// SIMATIC S7-200 project (STEP 7-Micro/WIN), CPU 224XP CN REL 02.01

SYMBOL_TABLE USUARIO1
C_1              VD100
C_0              VD110
y_k              VD180
r_k              VD190
u_k              VD120
xh1_k_1          VD130
xh1_k            VD140
xh2_k_1          VD300
xh2_k            VD160
xh3_k_1          VD170
xh3_k            VD200
xp1_k            VD210    // X1_v
xp2_k            VD220    // X2_v
xp3_k            VD230    // X3_v
Ao               VD310
Bo               VD320
Co               VD330
Do               VD340
Eo               VD350
Fo               VD360
Go               VD370
Ho               VD380
Io               VD390
Jo               VD400
L1o              VD410
L2o              VD420
L3o              VD430
e_k              VD270
Ee               VD240
r_k_1            VD250
u_k_1            VD150
k1o              VD440
k2o              VD450
k3o              VD460
END_SYMBOL_TABLE

ORGANIZATION_BLOCK PRINCIPAL:OB1
TITLE=COMENTARIOS DEL PROGRAMA
BEGIN
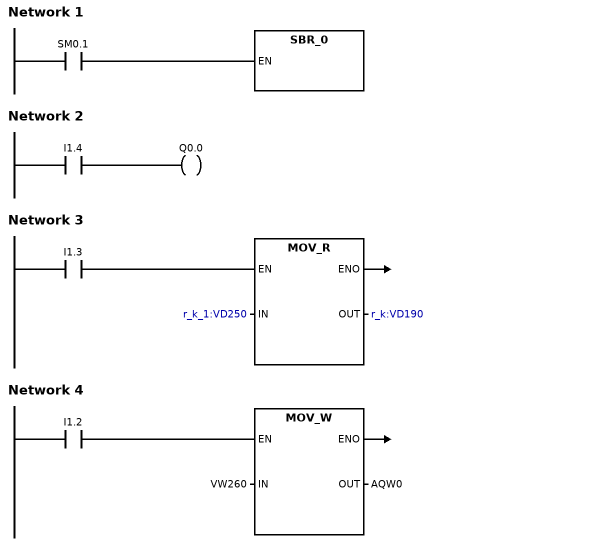
Network 1
LD     SM0.1
CALL   SBR_0:SBR0
Network 2
LD     I1.4
=      Q0.0
Network 3
LD     I1.3
MOVR   r_k_1:VD250, r_k:VD190
Network 4
LD     I1.2
MOVW   VW260, AQW0
END_ORGANIZATION_BLOCK

SUBROUTINE_BLOCK SBR_0:SBR0
TITLE=COMENTARIOS DE LA SUBRUTINA
BEGIN
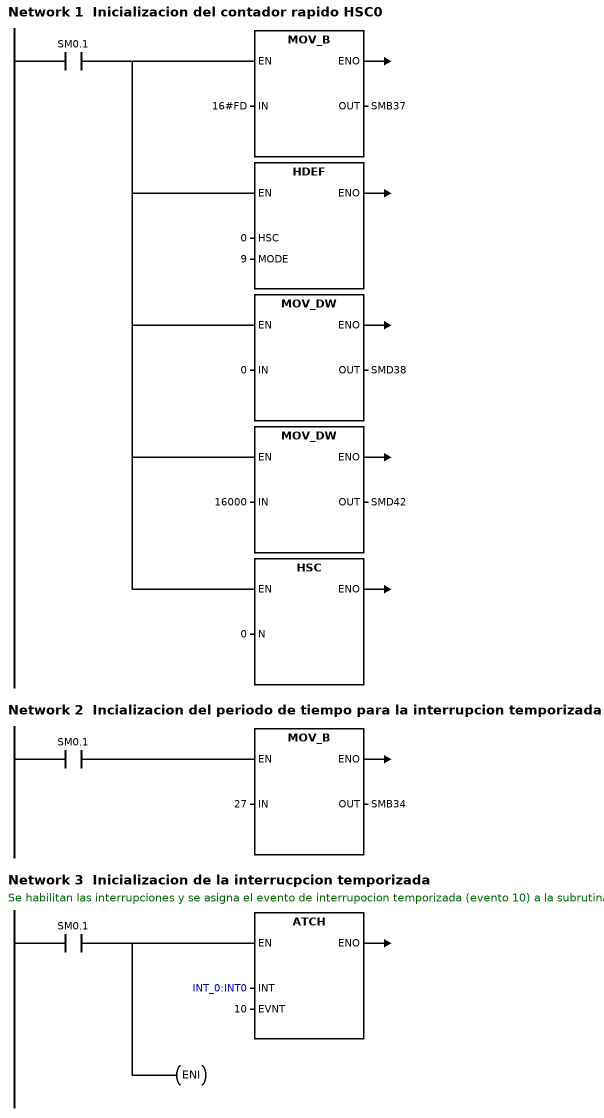
Network 1 // Inicializacion del contador rapido HSC0
LD     SM0.1
MOVB   16#FD, SMB37
HDEF   0, 9
MOVD   0, SMD38
MOVD   16000, SMD42
HSC    0
Network 2 // Incializacion del periodo de tiempo para la interrupcion temporizada
LD     SM0.1
MOVB   27, SMB34
Network 3 // Inicializacion de la interrucpcion temporizada
// Se habilitan las interrupciones y se asigna el evento de interrupocion temporizada (evento 10) a la subrutina de interrupcion INT_0
LD     SM0.1
ATCH   INT_0:INT0, 10
ENI
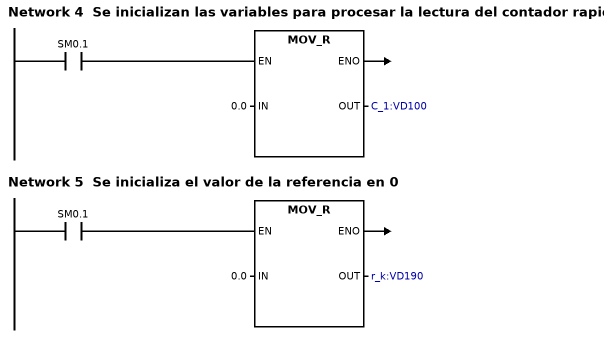
Network 4 // Se inicializan las variables para procesar la lectura del contador rapido HSC0
LD     SM0.1
MOVR   0.0, C_1:VD100
Network 5 // Se inicializa el valor de la referencia en 0
LD     SM0.1
MOVR   0.0, r_k:VD190
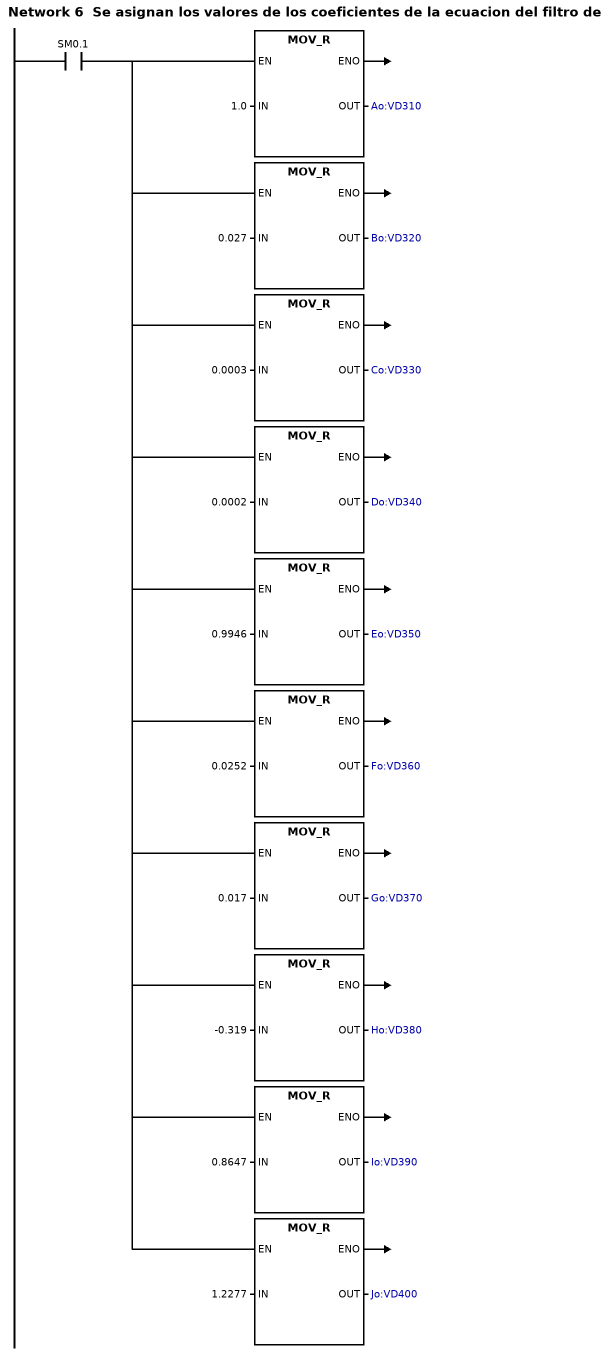
Network 6 // Se asignan los valores de los coeficientes de la ecuacion del filtro de KALMAN
LD     SM0.1
MOVR   1.0, Ao:VD310
MOVR   0.027, Bo:VD320
MOVR   0.0003, Co:VD330
MOVR   0.0002, Do:VD340
MOVR   0.9946, Eo:VD350
MOVR   0.0252, Fo:VD360
MOVR   0.017, Go:VD370
MOVR   -0.319, Ho:VD380
MOVR   0.8647, Io:VD390
MOVR   1.2277, Jo:VD400
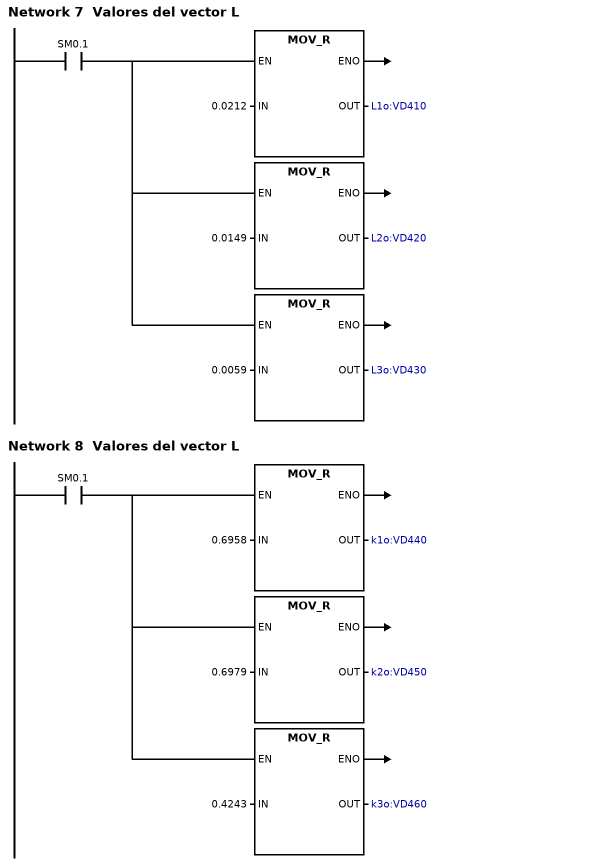
Network 7 // Valores del vector L
LD     SM0.1
MOVR   0.0212, L1o:VD410
MOVR   0.0149, L2o:VD420
MOVR   0.0059, L3o:VD430
Network 8 // Valores del vector L
LD     SM0.1
MOVR   0.6958, k1o:VD440
MOVR   0.6979, k2o:VD450
MOVR   0.4243, k3o:VD460
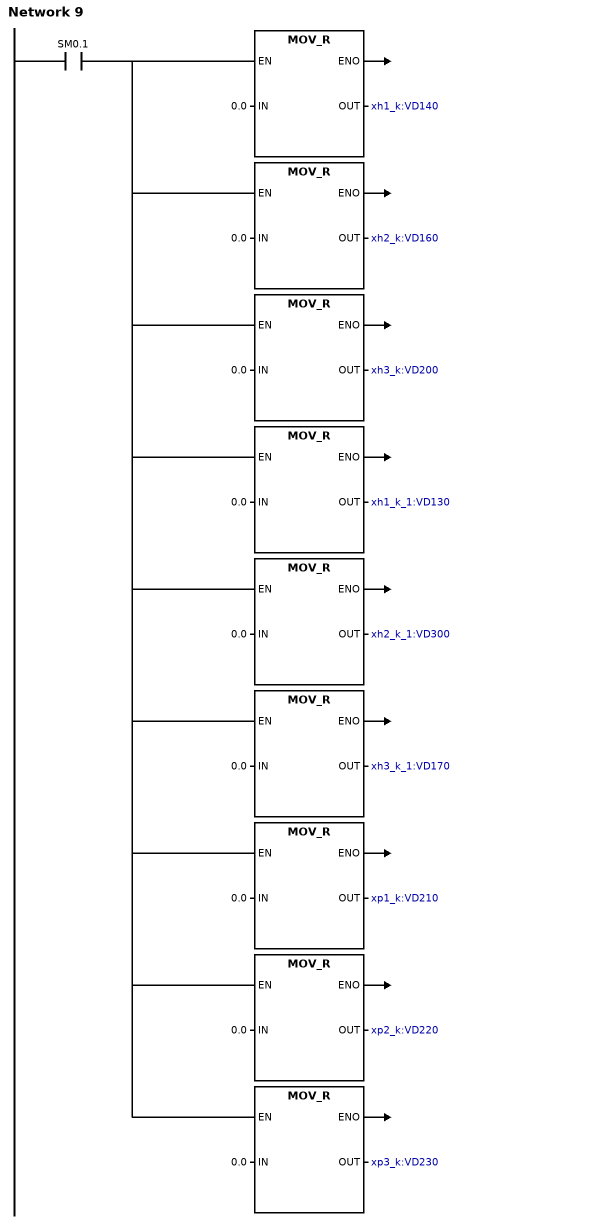
Network 9
LD     SM0.1
MOVR   0.0, xh1_k:VD140
MOVR   0.0, xh2_k:VD160
MOVR   0.0, xh3_k:VD200
MOVR   0.0, xh1_k_1:VD130
MOVR   0.0, xh2_k_1:VD300
MOVR   0.0, xh3_k_1:VD170
MOVR   0.0, xp1_k:VD210
MOVR   0.0, xp2_k:VD220
MOVR   0.0, xp3_k:VD230
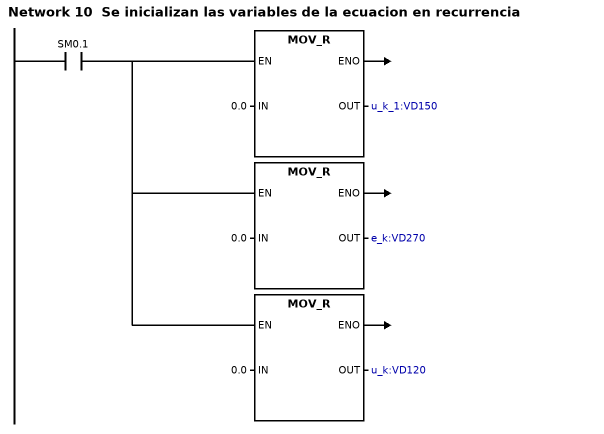
Network 10 // Se inicializan las variables de la ecuacion en recurrencia
LD     SM0.1
MOVR   0.0, u_k_1:VD150
MOVR   0.0, e_k:VD270
MOVR   0.0, u_k:VD120
END_SUBROUTINE_BLOCK

INTERRUPT_BLOCK INT_0:INT0
TITLE=COMENTARIOS DE LA RUTINA DE INTERRUPCIÓN
BEGIN
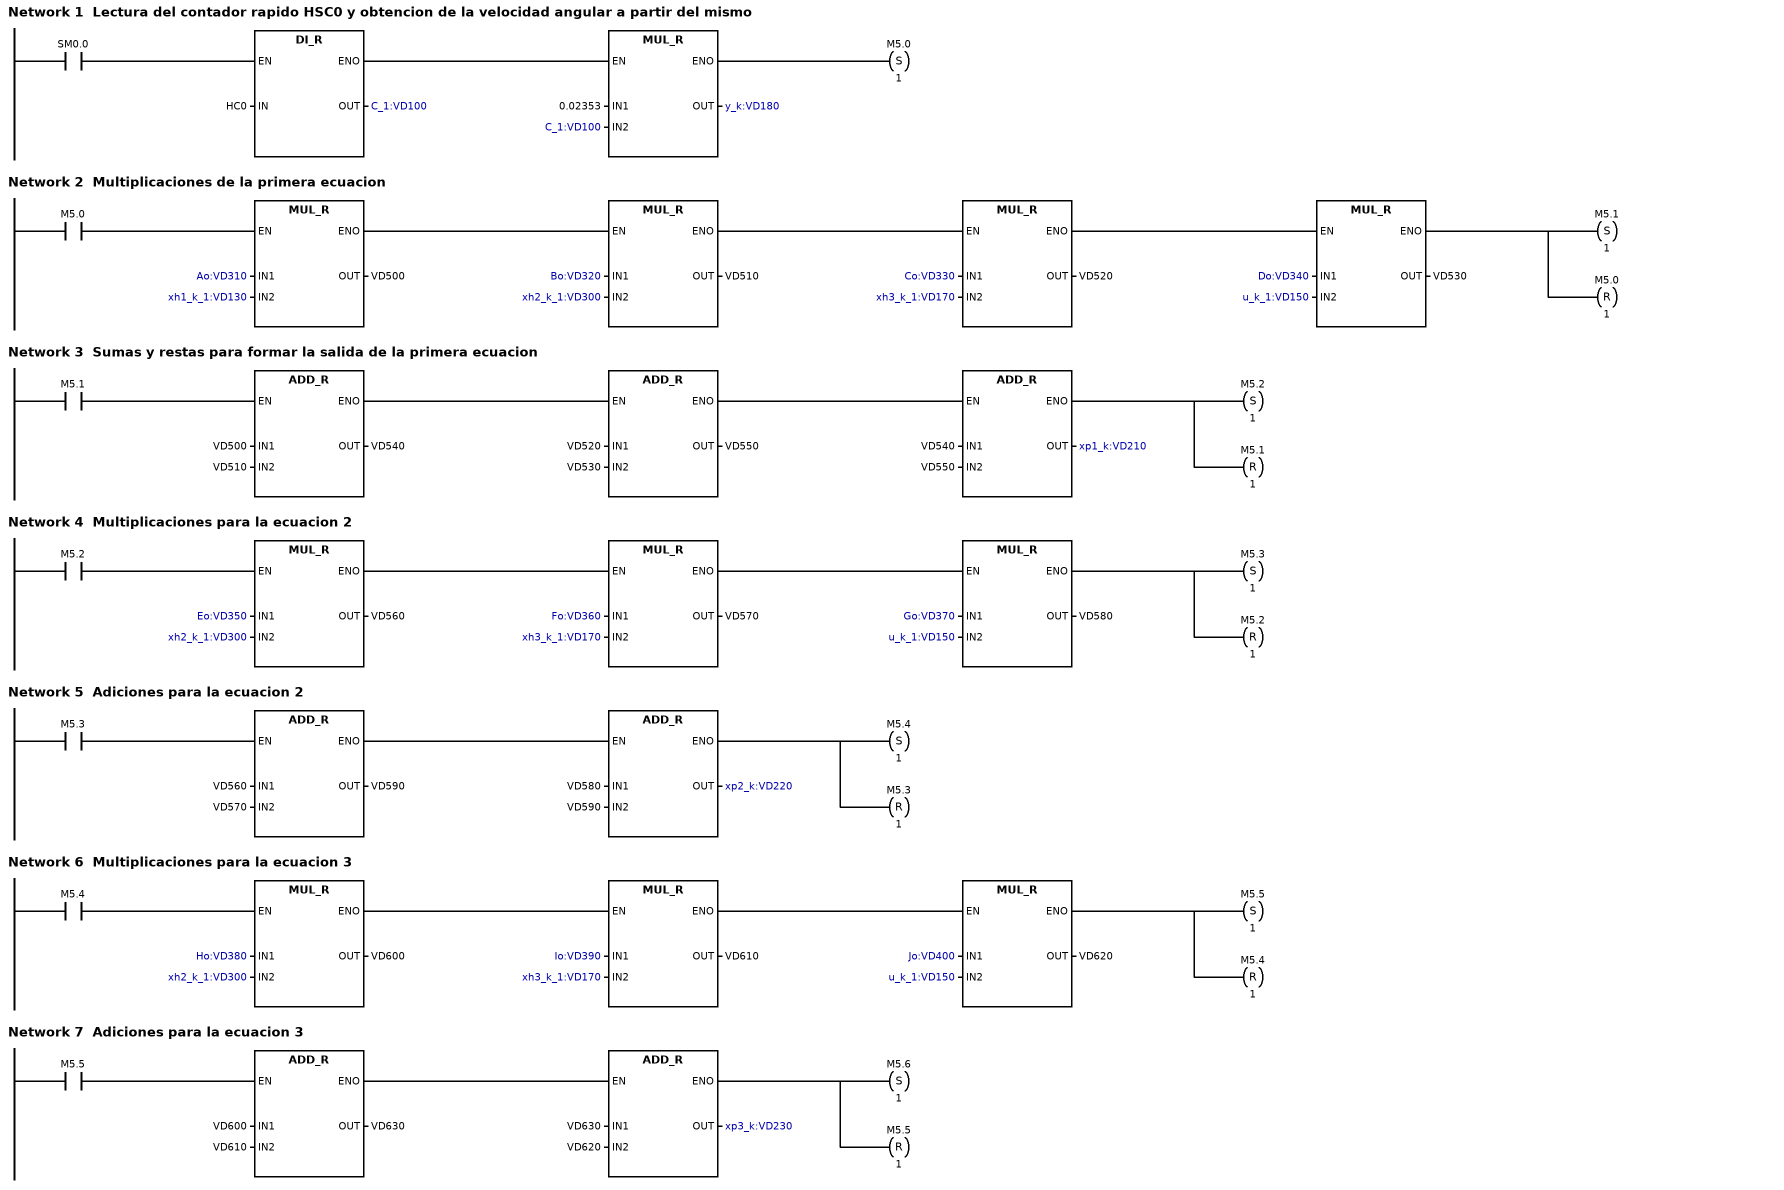
Network 1 // Lectura del contador rapido HSC0 y obtencion de la velocidad angular a partir del mismo
LD     SM0.0
DTR    HC0, C_1:VD100
AENO
MOVR   0.02353, y_k:VD180
AENO
*R     C_1:VD100, y_k:VD180
AENO
S      M5.0, 1
Network 2 // Multiplicaciones de la primera ecuacion 
LD     M5.0
MOVR   Ao:VD310, VD500
AENO
*R     xh1_k_1:VD130, VD500
AENO
MOVR   Bo:VD320, VD510
AENO
*R     xh2_k_1:VD300, VD510
AENO
MOVR   Co:VD330, VD520
AENO
*R     xh3_k_1:VD170, VD520
AENO
MOVR   Do:VD340, VD530
AENO
*R     u_k_1:VD150, VD530
AENO
S      M5.1, 1
R      M5.0, 1
Network 3 // Sumas y restas para formar la salida de la primera ecuacion
LD     M5.1
MOVR   VD500, VD540
AENO
+R     VD510, VD540
AENO
MOVR   VD520, VD550
AENO
+R     VD530, VD550
AENO
MOVR   VD540, xp1_k:VD210
AENO
+R     VD550, xp1_k:VD210
AENO
S      M5.2, 1
R      M5.1, 1
Network 4 // Multiplicaciones para la ecuacion 2
LD     M5.2
MOVR   Eo:VD350, VD560
AENO
*R     xh2_k_1:VD300, VD560
AENO
MOVR   Fo:VD360, VD570
AENO
*R     xh3_k_1:VD170, VD570
AENO
MOVR   Go:VD370, VD580
AENO
*R     u_k_1:VD150, VD580
AENO
S      M5.3, 1
R      M5.2, 1
Network 5 // Adiciones para la ecuacion 2
LD     M5.3
MOVR   VD560, VD590
AENO
+R     VD570, VD590
AENO
MOVR   VD580, xp2_k:VD220
AENO
+R     VD590, xp2_k:VD220
AENO
S      M5.4, 1
R      M5.3, 1
Network 6 // Multiplicaciones para la ecuacion 3
LD     M5.4
MOVR   Ho:VD380, VD600
AENO
*R     xh2_k_1:VD300, VD600
AENO
MOVR   Io:VD390, VD610
AENO
*R     xh3_k_1:VD170, VD610
AENO
MOVR   Jo:VD400, VD620
AENO
*R     u_k_1:VD150, VD620
AENO
S      M5.5, 1
R      M5.4, 1
Network 7 // Adiciones para la ecuacion 3
LD     M5.5
MOVR   VD600, VD630
AENO
+R     VD610, VD630
AENO
MOVR   VD630, xp3_k:VD230
AENO
+R     VD620, xp3_k:VD230
AENO
S      M5.6, 1
R      M5.5, 1
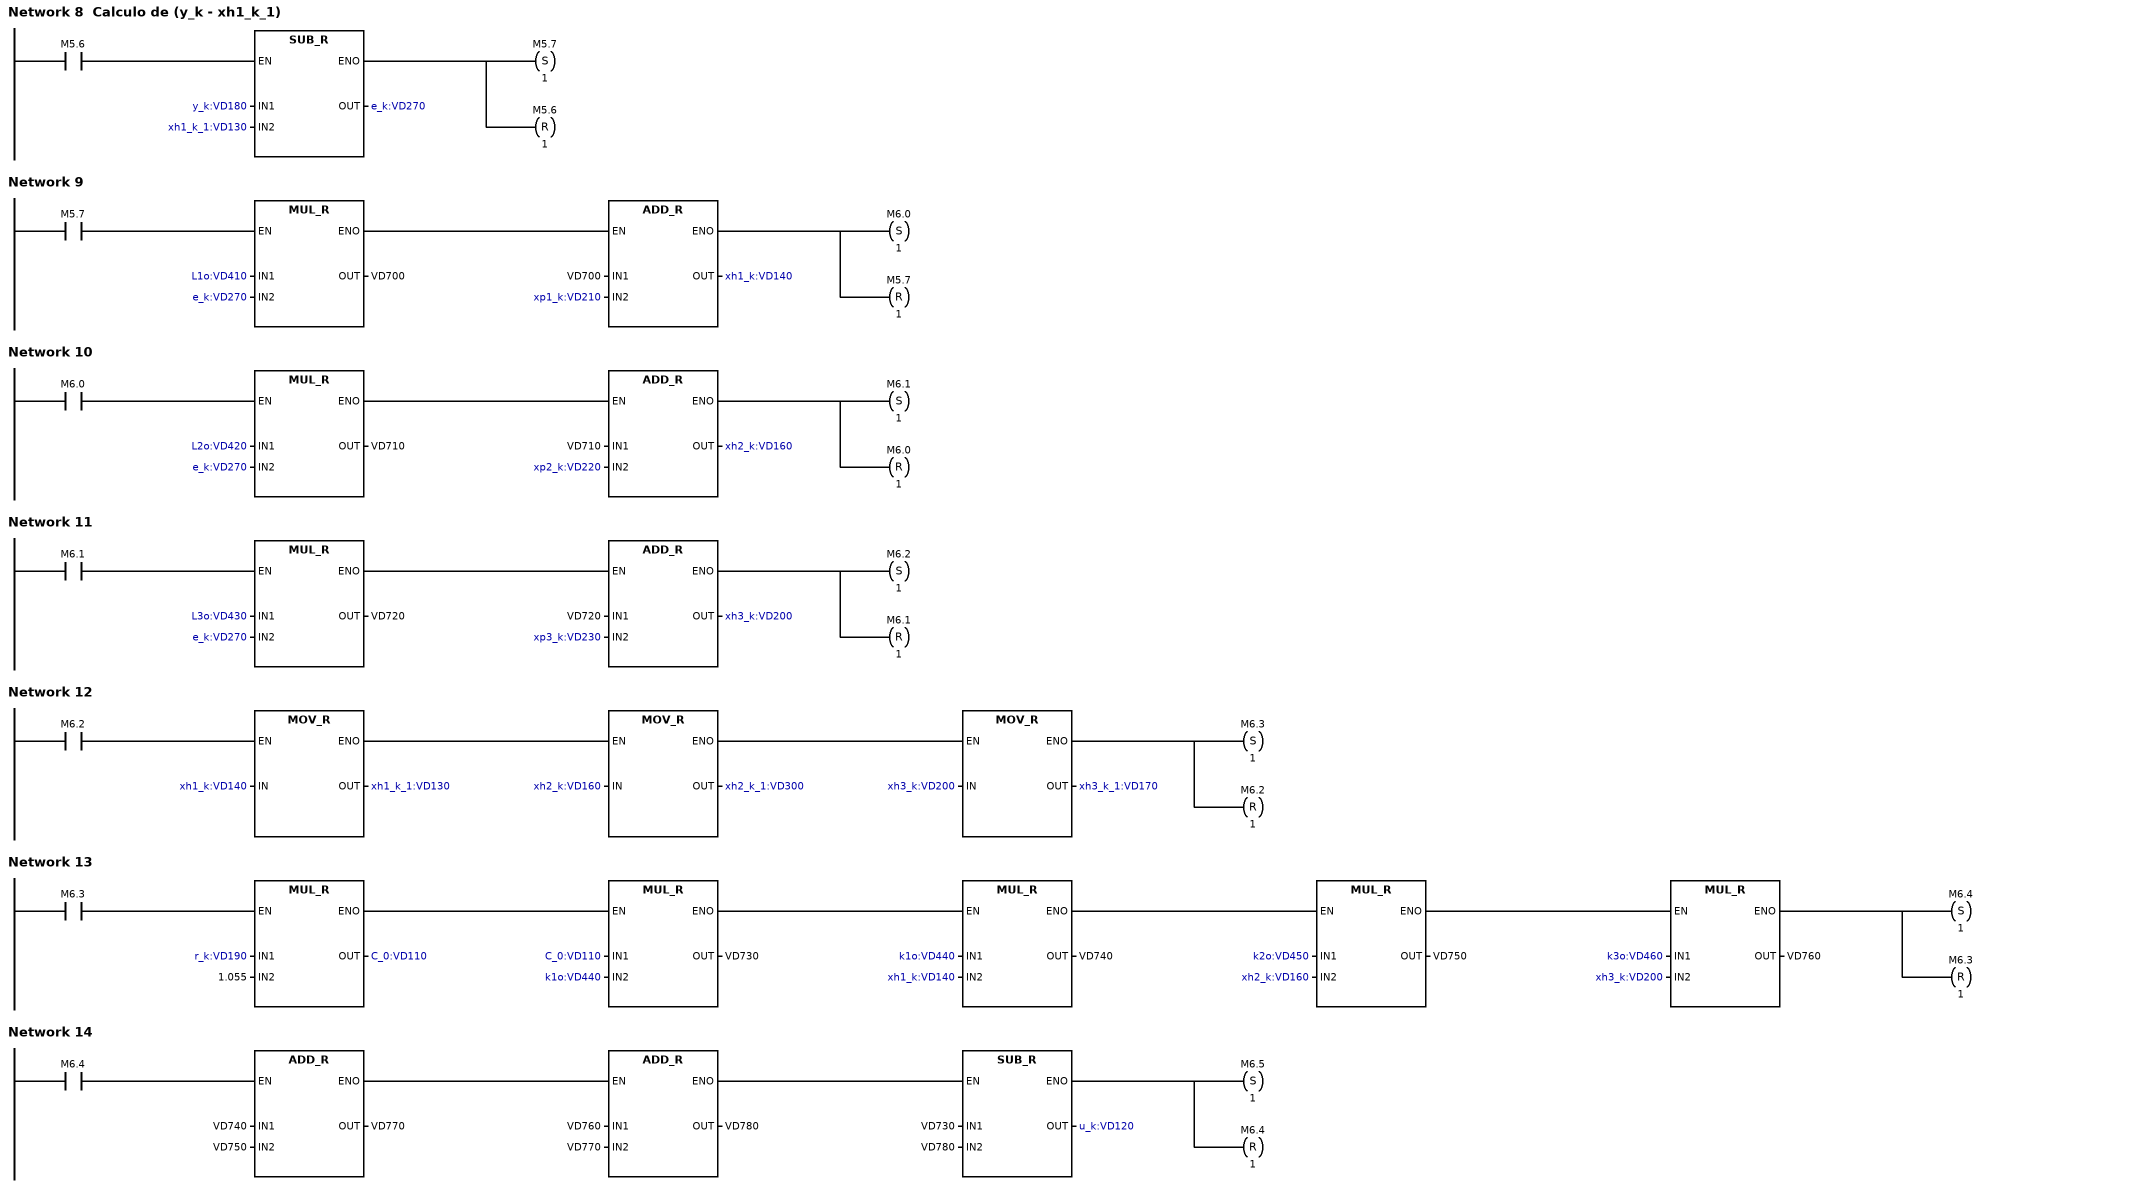
Network 8 // Calculo de (y_k - xh1_k_1)
LD     M5.6
MOVR   y_k:VD180, e_k:VD270
AENO
-R     xh1_k_1:VD130, e_k:VD270
AENO
S      M5.7, 1
R      M5.6, 1
Network 9
LD     M5.7
MOVR   L1o:VD410, VD700
AENO
*R     e_k:VD270, VD700
AENO
MOVR   VD700, xh1_k:VD140
AENO
+R     xp1_k:VD210, xh1_k:VD140
AENO
S      M6.0, 1
R      M5.7, 1
Network 10
LD     M6.0
MOVR   L2o:VD420, VD710
AENO
*R     e_k:VD270, VD710
AENO
MOVR   VD710, xh2_k:VD160
AENO
+R     xp2_k:VD220, xh2_k:VD160
AENO
S      M6.1, 1
R      M6.0, 1
Network 11
LD     M6.1
MOVR   L3o:VD430, VD720
AENO
*R     e_k:VD270, VD720
AENO
MOVR   VD720, xh3_k:VD200
AENO
+R     xp3_k:VD230, xh3_k:VD200
AENO
S      M6.2, 1
R      M6.1, 1
Network 12
LD     M6.2
MOVR   xh1_k:VD140, xh1_k_1:VD130
AENO
MOVR   xh2_k:VD160, xh2_k_1:VD300
AENO
MOVR   xh3_k:VD200, xh3_k_1:VD170
AENO
S      M6.3, 1
R      M6.2, 1
Network 13
LD     M6.3
MOVR   r_k:VD190, C_0:VD110
AENO
*R     1.055, C_0:VD110
AENO
MOVR   C_0:VD110, VD730
AENO
*R     k1o:VD440, VD730
AENO
MOVR   k1o:VD440, VD740
AENO
*R     xh1_k:VD140, VD740
AENO
MOVR   k2o:VD450, VD750
AENO
*R     xh2_k:VD160, VD750
AENO
MOVR   k3o:VD460, VD760
AENO
*R     xh3_k:VD200, VD760
AENO
S      M6.4, 1
R      M6.3, 1
Network 14
LD     M6.4
MOVR   VD740, VD770
AENO
+R     VD750, VD770
AENO
MOVR   VD760, VD780
AENO
+R     VD770, VD780
AENO
MOVR   VD730, u_k:VD120
AENO
-R     VD780, u_k:VD120
AENO
S      M6.5, 1
R      M6.4, 1
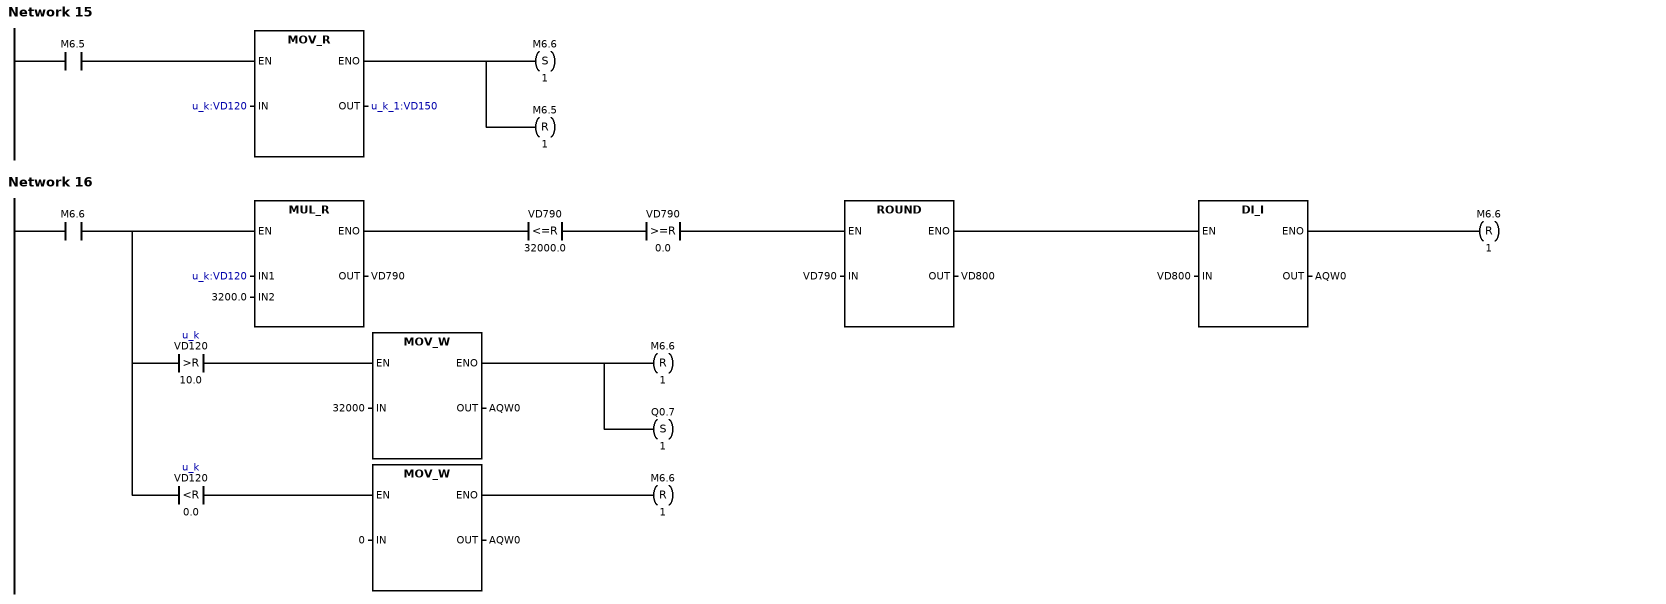
Network 15
LD     M6.5
MOVR   u_k:VD120, u_k_1:VD150
AENO
S      M6.6, 1
R      M6.5, 1
Network 16
LD     M6.6
LPS
MOVR   u_k:VD120, VD790
AENO
*R     3200.0, VD790
AENO
AR<=   VD790, 32000.0
AR>=   VD790, 0.0
ROUND  VD790, VD800
AENO
DTI    VD800, AQW0
AENO
R      M6.6, 1
LRD
AR>    u_k:VD120, 10.0
MOVW   32000, AQW0
AENO
R      M6.6, 1
S      Q0.7, 1
LPP
AR<    u_k:VD120, 0.0
MOVW   0, AQW0
AENO
R      M6.6, 1
END_INTERRUPT_BLOCK
